// TwinCAT 3 PLC project PLC
// libraries:
//   Tc2_Standard, * (Beckhoff Automation GmbH)
// project tree:
//   DUTs/ E_State.TcDUT
//   duts/ e_state.TcDUT
//   GVLs/Old/ GVL_Moved.TcGVL (not stored)
//   / PlcTask.TcTTO
//   POUs/ FB_Gone.TcPOU (not stored), fb_listed.TcPOU, MAIN.TcPOU, MAIN.TcPOU

CONFIGURATION PLC
    RESOURCE PLC ON TwinCAT3
        TASK PlcTask(INTERVAL := ?, PRIORITY := 0);
    END_RESOURCE
END_CONFIGURATION

// ---- DUTs/E_State.TcDUT
TYPE E_State :
(
  Idle,
  Busy
);
END_TYPE

// ---- duts/e_state.TcDUT
TYPE E_State :
(
  Idle,
  Busy
);
END_TYPE

// ---- POUs/fb_listed.TcPOU
FUNCTION_BLOCK FB_Listed

END_FUNCTION_BLOCK

// ---- POUs/MAIN.TcPOU
PROGRAM MAIN

END_PROGRAM

// ---- POUs/MAIN.TcPOU
PROGRAM MAIN

END_PROGRAM
